// TIA Portal V20 export
// export: Created 2026-10-20T18:55:21.550557Z, ExportSetting None, DisplayName Totally Integrated Automation Portal, DisplayVersion V20 Update 6, DisplayName TIA Portal Openness, DisplayVersion V20 Update 6, DisplayName TIA Portal Version Control Interface, DisplayVersion V20 Update 6, DisplayName SINAMICS Startdrive Advanced, DisplayVersion V20 SP1, DisplayName SINAMICS Startdrive G130, G150, S120, S150, SINAMICS MV, G220, S200, S210, DisplayVersion V20 SP1, DisplayName SINAMICS Startdrive G110M, G120, G120C, G120D, G120P, G115D, DisplayVersion V20 SP1, DisplayName STEP 7 Professional, DisplayVersion V20 Update 6, DisplayName STEP 7 Safety, DisplayVersion V20 Update 2, DisplayName WinCC Basic/Comfort/Advanced, DisplayVersion V20 Update 6, DisplayName WinCC Unified, DisplayVersion V20 Update 6
VAR_GLOBAL   // PLC tag table "IO_Encoders_4"
   "LE_Warnings(4)" AT %IW1195 : Int;
   "LE_Speed(4)" AT %IW1193 : Int;   // 0 ...65535
   "LE_Status(4)" AT %IW1187 : UInt;
   "LE_X_Unsafe_Position(4)" AT %ID1189 : DInt;
   "AE_Status_1(4)" AT %IW1281 : UInt;   // 8 … 0 - Reserved / 9 - Control requested / 11,10 - Reserved / 15...12 - Encoder’s Sign-of-Life (not relevant)
   "AE_Control_Word_2(4)" AT %QW1058 : UInt;   // 10 … 0 - Reserved / 11 - Preset mode / 12 - Activate preset value / 13 - Request for the absolute position value / 14 - Activate park mode / 15 - Acknowledging a sensor error
   "AE_Status_2(4)" AT %IW1283 : UInt;   // 9 … 0 - Not supported / 10 - Reserved / 11 - Requirement of error acknowledgement detected / 12 - Status of the Preset function (set/shift of home position executed) / 13 - Transmission of absolute position value / 14 - Park mode activated / 15 - Encoder error
   "AE_Position_2(4)" AT %ID1289 : DInt;
   "AE_Position_1(4)" AT %ID1285 : DInt;
   "AE_Speed(4)" AT %IW1293 : Int;
   "AE_Control_Word_1(4)" AT %QW1056 : UInt;   // 11, 9, 8, 6 … 0 - Reserved / 7 - Fault acknowledge / 10 - Control by PLC / 15...12 - Master’s Sign-of-Life (not relevant)
END_VAR
